(* IEC 61131-3 sources: plc-st-coding-agent/progress/evidence/f14_v5_public_pilot_20261112/jobs/codex_minimax-m27, 24 files *)

(* ---- public-easy-01.candidate_01.st ---- *)
(*
ENGINEERING_CONTRACT - Filling Line Control FB
==============================================
State Machine: Sequential, 6 states (IDLE→CLEANING→FILLING→CAPPING→PACKING→COMPLETED→IDLE)
---------------------------------------------------------------------------------
| State       | Activation         | Retention              | Reset/Deactivation            |
---------------------------------------------------------------------------------
| IDLE        | bottleSensor=TRUE  | Hold until bottle      | Deact on bottleSensor:=TRUE   |
| CLEANING    | cleaningConfirm    | Pump_Motor ON hold     | Deact on cleaningConfirm      |
| FILLING     | fillingConfirm     | Filling_Valve ON hold  | Deact on fillingConfirm       |
| CAPPING     | cappingConfirm     | Capping_Machine ON hold| Deact on cappingConfirm       |
| PACKING     | packingConfirm     | Packing_Machine ON hold| Deact on packingConfirm       |
| COMPLETED   | packingConfirm     | Completion_Light ON    | Deact on finishedButton       |
---------------------------------------------------------------------------------
Priority: IDLE > COMPLETED > CLEANING > FILLING > CAPPING > PACKING (same-scan)
Units: All inputs/outputs BOOL; all states enumerated; no TIME/LTIME used
Boundaries: bottleSensor triggers only from IDLE; finishedButton resets only from COMPLETED
PUB refs: PUB001, PUB003, PUB004, PUB005, PUB006, PUB007, PUB008
---------------------------------------------------------------------------------
*)
FUNCTION_BLOCK FillingLineControl
VAR
    eState : EFillState := EFillState.IDLE;
END_VAR

TYPE EFillState :
(
    IDLE       := 0,
    CLEANING   := 1,
    FILLING    := 2,
    CAPPING    := 3,
    PACKING    := 4,
    COMPLETED  := 5
);
END_TYPE;

CASE eState OF
    EFillState.IDLE:
        Pump_Motor       := FALSE;
        Filling_Valve    := FALSE;
        Capping_Machine  := FALSE;
        Packing_Machine  := FALSE;
        Completion_Light := FALSE;

        IF bottleSensor THEN
            eState := EFillState.CLEANING;
        END_IF;

    EFillState.CLEANING:
        Pump_Motor       := TRUE;
        Filling_Valve    := FALSE;
        Capping_Machine  := FALSE;
        Packing_Machine  := FALSE;
        Completion_Light := FALSE;

        IF cleaningConfirmButton THEN
            eState := EFillState.FILLING;
        END_IF;

    EFillState.FILLING:
        Pump_Motor       := TRUE;
        Filling_Valve    := TRUE;
        Capping_Machine  := FALSE;
        Packing_Machine  := FALSE;
        Completion_Light := FALSE;

        IF fillingConfirmButton THEN
            eState := EFillState.CAPPING;
        END_IF;

    EFillState.CAPPING:
        Pump_Motor       := TRUE;
        Filling_Valve    := FALSE;
        Capping_Machine  := TRUE;
        Packing_Machine  := FALSE;
        Completion_Light := FALSE;

        IF cappingConfirmButton THEN
            eState := EFillState.PACKING;
        END_IF;

    EFillState.PACKING:
        Pump_Motor       := TRUE;
        Filling_Valve    := FALSE;
        Capping_Machine  := FALSE;
        Packing_Machine  := TRUE;
        Completion_Light := FALSE;

        IF packingConfirmButton THEN
            eState := EFillState.COMPLETED;
        END_IF;

    EFillState.COMPLETED:
        Pump_Motor       := TRUE;
        Filling_Valve    := FALSE;
        Capping_Machine  := FALSE;
        Packing_Machine  := FALSE;
        Completion_Light := TRUE;

        IF finishedButton THEN
            eState := EFillState.IDLE;
        END_IF;

END_CASE;

END_FUNCTION_BLOCK

(* ---- public-easy-01.candidate_02.st ---- *)
(*
ENGINEERING_CONTRACT - Filling Line Control FB
==============================================
State Machine: Sequential, 6 states (IDLE→CLEANING→FILLING→CAPPING→PACKING→COMPLETED→IDLE)
---------------------------------------------------------------------------------
| State       | Activation         | Retention              | Reset/Deactivation            |
---------------------------------------------------------------------------------
| IDLE        | bottleSensor=TRUE  | Hold until bottle      | Deact on bottleSensor:=TRUE   |
| CLEANING    | cleaningConfirm    | Pump_Motor ON hold     | Deact on cleaningConfirm      |
| FILLING     | fillingConfirm     | Filling_Valve ON hold  | Deact on fillingConfirm       |
| CAPPING     | cappingConfirm     | Capping_Machine ON hold| Deact on cappingConfirm       |
| PACKING     | packingConfirm     | Packing_Machine ON hold| Deact on packingConfirm       |
| COMPLETED   | packingConfirm     | Completion_Light ON    | Deact on finishedButton       |
---------------------------------------------------------------------------------
Priority: IDLE > COMPLETED > CLEANING > FILLING > CAPPING > PACKING (same-scan)
Units: All inputs/outputs BOOL; all states enumerated; no TIME/LTIME used
Boundaries: bottleSensor triggers only from IDLE; finishedButton resets only from COMPLETED
PUB refs: PUB001, PUB003, PUB004, PUB005, PUB006, PUB007, PUB008
---------------------------------------------------------------------------------
*)
TYPE EFillState :
(
    IDLE       := 0,
    CLEANING   := 1,
    FILLING    := 2,
    CAPPING    := 3,
    PACKING    := 4,
    COMPLETED  := 5
);
END_TYPE;

FUNCTION_BLOCK FillingLineControl
VAR_INPUT
    bottleSensor           : BOOL;
    cleaningConfirmButton  : BOOL;
    fillingConfirmButton   : BOOL;
    cappingConfirmButton   : BOOL;
    packingConfirmButton   : BOOL;
    finishedButton         : BOOL;
END_VAR
VAR_OUTPUT
    Pump_Motor       : BOOL;
    Filling_Valve    : BOOL;
    Capping_Machine  : BOOL;
    Packing_Machine  : BOOL;
    Completion_Light : BOOL;
END_VAR
VAR
    eState : EFillState := EFillState.IDLE;
END_VAR

CASE eState OF
    EFillState.IDLE:
        Pump_Motor       := FALSE;
        Filling_Valve    := FALSE;
        Capping_Machine  := FALSE;
        Packing_Machine  := FALSE;
        Completion_Light := FALSE;

        IF bottleSensor THEN
            eState := EFillState.CLEANING;
        END_IF;

    EFillState.CLEANING:
        Pump_Motor       := TRUE;
        Filling_Valve    := FALSE;
        Capping_Machine  := FALSE;
        Packing_Machine  := FALSE;
        Completion_Light := FALSE;

        IF cleaningConfirmButton THEN
            eState := EFillState.FILLING;
        END_IF;

    EFillState.FILLING:
        Pump_Motor       := FALSE;
        Filling_Valve    := TRUE;
        Capping_Machine  := FALSE;
        Packing_Machine  := FALSE;
        Completion_Light := FALSE;

        IF fillingConfirmButton THEN
            eState := EFillState.CAPPING;
        END_IF;

    EFillState.CAPPING:
        Pump_Motor       := FALSE;
        Filling_Valve    := FALSE;
        Capping_Machine  := TRUE;
        Packing_Machine  := FALSE;
        Completion_Light := FALSE;

        IF cappingConfirmButton THEN
            eState := EFillState.PACKING;
        END_IF;

    EFillState.PACKING:
        Pump_Motor       := FALSE;
        Filling_Valve    := FALSE;
        Capping_Machine  := FALSE;
        Packing_Machine  := TRUE;
        Completion_Light := FALSE;

        IF packingConfirmButton THEN
            eState := EFillState.COMPLETED;
        END_IF;

    EFillState.COMPLETED:
        Pump_Motor       := FALSE;
        Filling_Valve    := FALSE;
        Capping_Machine  := FALSE;
        Packing_Machine  := FALSE;
        Completion_Light := TRUE;

        IF finishedButton THEN
            eState := EFillState.IDLE;
        END_IF;

END_CASE;

END_FUNCTION_BLOCK

(* ---- public-easy-01.raw_candidate_01.st ---- *)
(*
ENGINEERING_CONTRACT - Filling Line Control FB
==============================================
State Machine: Sequential, 6 states (IDLE→CLEANING→FILLING→CAPPING→PACKING→COMPLETED→IDLE)
---------------------------------------------------------------------------------
| State       | Activation         | Retention              | Reset/Deactivation            |
---------------------------------------------------------------------------------
| IDLE        | bottleSensor=TRUE  | Hold until bottle      | Deact on bottleSensor:=TRUE   |
| CLEANING    | cleaningConfirm    | Pump_Motor ON hold     | Deact on cleaningConfirm      |
| FILLING     | fillingConfirm     | Filling_Valve ON hold  | Deact on fillingConfirm       |
| CAPPING     | cappingConfirm     | Capping_Machine ON hold| Deact on cappingConfirm       |
| PACKING     | packingConfirm     | Packing_Machine ON hold| Deact on packingConfirm       |
| COMPLETED   | packingConfirm     | Completion_Light ON    | Deact on finishedButton       |
---------------------------------------------------------------------------------
Priority: IDLE > COMPLETED > CLEANING > FILLING > CAPPING > PACKING (same-scan)
Units: All inputs/outputs BOOL; all states enumerated; no TIME/LTIME used
Boundaries: bottleSensor triggers only from IDLE; finishedButton resets only from COMPLETED
PUB refs: PUB001, PUB003, PUB004, PUB005, PUB006, PUB007, PUB008
---------------------------------------------------------------------------------
*)
FUNCTION_BLOCK FillingLineControl
VAR
    eState : EFillState := EFillState.IDLE;
END_VAR

TYPE EFillState :
(
    IDLE       := 0,
    CLEANING   := 1,
    FILLING    := 2,
    CAPPING    := 3,
    PACKING    := 4,
    COMPLETED  := 5
);
END_TYPE

CASE eState OF
    EFillState.IDLE:
        Pump_Motor       := FALSE;
        Filling_Valve    := FALSE;
        Capping_Machine  := FALSE;
        Packing_Machine  := FALSE;
        Completion_Light := FALSE;

        IF bottleSensor THEN
            eState := EFillState.CLEANING;
        END_IF;

    EFillState.CLEANING:
        Pump_Motor       := TRUE;
        Filling_Valve    := FALSE;
        Capping_Machine  := FALSE;
        Packing_Machine  := FALSE;
        Completion_Light := FALSE;

        IF cleaningConfirmButton THEN
            eState := EFillState.FILLING;
        END_IF;

    EFillState.FILLING:
        Pump_Motor       := TRUE;
        Filling_Valve    := TRUE;
        Capping_Machine  := FALSE;
        Packing_Machine  := FALSE;
        Completion_Light := FALSE;

        IF fillingConfirmButton THEN
            eState := EFillState.CAPPING;
        END_IF;

    EFillState.CAPPING:
        Pump_Motor       := TRUE;
        Filling_Valve    := FALSE;
        Capping_Machine  := TRUE;
        Packing_Machine  := FALSE;
        Completion_Light := FALSE;

        IF cappingConfirmButton THEN
            eState := EFillState.PACKING;
        END_IF;

    EFillState.PACKING:
        Pump_Motor       := TRUE;
        Filling_Valve    := FALSE;
        Capping_Machine  := FALSE;
        Packing_Machine  := TRUE;
        Completion_Light := FALSE;

        IF packingConfirmButton THEN
            eState := EFillState.COMPLETED;
        END_IF;

    EFillState.COMPLETED:
        Pump_Motor       := TRUE;
        Filling_Valve    := FALSE;
        Capping_Machine  := FALSE;
        Packing_Machine  := FALSE;
        Completion_Light := TRUE;

        IF finishedButton THEN
            eState := EFillState.IDLE;
        END_IF;

END_CASE;

END_FUNCTION_BLOCK

(* ---- public-easy-01.raw_candidate_02.st ---- *)
(*
ENGINEERING_CONTRACT - Filling Line Control FB
==============================================
State Machine: Sequential, 6 states (IDLE→CLEANING→FILLING→CAPPING→PACKING→COMPLETED→IDLE)
---------------------------------------------------------------------------------
| State       | Activation         | Retention              | Reset/Deactivation            |
---------------------------------------------------------------------------------
| IDLE        | bottleSensor=TRUE  | Hold until bottle      | Deact on bottleSensor:=TRUE   |
| CLEANING    | cleaningConfirm    | Pump_Motor ON hold     | Deact on cleaningConfirm      |
| FILLING     | fillingConfirm     | Filling_Valve ON hold  | Deact on fillingConfirm       |
| CAPPING     | cappingConfirm     | Capping_Machine ON hold| Deact on cappingConfirm       |
| PACKING     | packingConfirm     | Packing_Machine ON hold| Deact on packingConfirm       |
| COMPLETED   | packingConfirm     | Completion_Light ON    | Deact on finishedButton       |
---------------------------------------------------------------------------------
Priority: IDLE > COMPLETED > CLEANING > FILLING > CAPPING > PACKING (same-scan)
Units: All inputs/outputs BOOL; all states enumerated; no TIME/LTIME used
Boundaries: bottleSensor triggers only from IDLE; finishedButton resets only from COMPLETED
PUB refs: PUB001, PUB003, PUB004, PUB005, PUB006, PUB007, PUB008
---------------------------------------------------------------------------------
*)
TYPE EFillState :
(
    IDLE       := 0,
    CLEANING   := 1,
    FILLING    := 2,
    CAPPING    := 3,
    PACKING    := 4,
    COMPLETED  := 5
);
END_TYPE

FUNCTION_BLOCK FillingLineControl
VAR_INPUT
    bottleSensor           : BOOL;
    cleaningConfirmButton  : BOOL;
    fillingConfirmButton   : BOOL;
    cappingConfirmButton   : BOOL;
    packingConfirmButton   : BOOL;
    finishedButton         : BOOL;
END_VAR
VAR_OUTPUT
    Pump_Motor       : BOOL;
    Filling_Valve    : BOOL;
    Capping_Machine  : BOOL;
    Packing_Machine  : BOOL;
    Completion_Light : BOOL;
END_VAR
VAR
    eState : EFillState := EFillState.IDLE;
END_VAR

CASE eState OF
    EFillState.IDLE:
        Pump_Motor       := FALSE;
        Filling_Valve    := FALSE;
        Capping_Machine  := FALSE;
        Packing_Machine  := FALSE;
        Completion_Light := FALSE;

        IF bottleSensor THEN
            eState := EFillState.CLEANING;
        END_IF;

    EFillState.CLEANING:
        Pump_Motor       := TRUE;
        Filling_Valve    := FALSE;
        Capping_Machine  := FALSE;
        Packing_Machine  := FALSE;
        Completion_Light := FALSE;

        IF cleaningConfirmButton THEN
            eState := EFillState.FILLING;
        END_IF;

    EFillState.FILLING:
        Pump_Motor       := FALSE;
        Filling_Valve    := TRUE;
        Capping_Machine  := FALSE;
        Packing_Machine  := FALSE;
        Completion_Light := FALSE;

        IF fillingConfirmButton THEN
            eState := EFillState.CAPPING;
        END_IF;

    EFillState.CAPPING:
        Pump_Motor       := FALSE;
        Filling_Valve    := FALSE;
        Capping_Machine  := TRUE;
        Packing_Machine  := FALSE;
        Completion_Light := FALSE;

        IF cappingConfirmButton THEN
            eState := EFillState.PACKING;
        END_IF;

    EFillState.PACKING:
        Pump_Motor       := FALSE;
        Filling_Valve    := FALSE;
        Capping_Machine  := FALSE;
        Packing_Machine  := TRUE;
        Completion_Light := FALSE;

        IF packingConfirmButton THEN
            eState := EFillState.COMPLETED;
        END_IF;

    EFillState.COMPLETED:
        Pump_Motor       := FALSE;
        Filling_Valve    := FALSE;
        Capping_Machine  := FALSE;
        Packing_Machine  := FALSE;
        Completion_Light := TRUE;

        IF finishedButton THEN
            eState := EFillState.IDLE;
        END_IF;

END_CASE;

END_FUNCTION_BLOCK

(* ---- public-easy-04.candidate_01.st ---- *)
FUNCTION_BLOCK JamPumpControl
VAR_INPUT
    VISCOSITY_OK    : BOOL;
    PASTE_E_STOP_NC : BOOL;
    DebounceTime    : TIME;
    CycleTime       : TIME;
END_VAR
VAR_OUTPUT
    VFD_RUN          : BOOL := FALSE;
    PUMP_MAINT_DUE   : BOOL := FALSE;
    PUMP_RUNTIME_ACC : LTIME := LTIME#0s;
END_VAR
VAR
    ViscosityDebounceTimer : TON;
    ViscosityDebounceAccum : LTIME := LTIME#0s;
    ViscosityValid         : BOOL := FALSE;
END_VAR
// ENGINEERING_CONTRACT
// | Output/State    | Activation         | Retention          | Reset/Deactivation                      | Priority | Units/Boundaries |
// |-----------------|--------------------|--------------------|-----------------------------------------|----------|-------------------|
// | VFD_RUN         | TRUE when safety   | Retained while     | Cleared on E-Stop or viscosity invalid  | Safety   | Boolean permissive|
// |                 | permissive AND     | conditions met     | (PUB003)                                | first    |                   |
// |                 | viscosity valid    |                    |                                         |          |                   |
// | PUMP_MAINT_DUE  | Set when runtime   | Latched TRUE       | No reset (informational only, PUB004)   | None     | 500h threshold    |
// |                 | >= 500h (PUB004)   |                    |                                         |          |                   |
// | PUMP_RUNTIME_ACC| Increments by      | Preserved when     | Init to 0 at power-up only (PUB005)     | None     | LTIME (nanoseconds)|
// |                 | CycleTime when     | VFD_RUN = FALSE    |                                         |          | 0 to max          |
// |                 | VFD_RUN = TRUE     | (PUB003)           |                                         |          |                   |
// |                 | (PUB003)          |                    |                                         |          |                   |
// | ViscosityValid  | After DebounceTime | Retained while     | Immediate on VISCITY_OK=FALSE or        | None     | Debounced state   |
// |                 | continuous TRUE    | VISCOSITY_OK=TRUE  | E-Stop (PUB002, PUB003)                 |          |                   |
// |                 | (PUB002)          | (PUB002)           |                                         |          |                   |
// | ViscosityDebounceAccum | Accumulates  | Reset to 0 when   | Reset on VISCOSITY_OK=FALSE or          | None     | LTIME nanoseconds |
// |                 | elapsed time when  | VISCOSITY_OK=FALSE | E-Stop (PUB003)                         |          | >= 0              |
// |                 | VISCOSITY_OK=TRUE  |                    |                                         |          |                   |

// Viscosity debouncing (PUB002)
IF NOT VISCOSITY_OK THEN
    ViscosityDebounceAccum := LTIME#0s;
    ViscosityValid := FALSE;
    ViscosityDebounceTimer(IN := FALSE);
ELSIF ViscosityValid THEN
    ViscosityDebounceTimer(IN := TRUE, PT := DebounceTime);
ELSE
    ViscosityDebounceAccum := ViscosityDebounceAccum + CycleTime;
    IF ViscosityDebounceAccum >= DebounceTime THEN
        ViscosityValid := TRUE;
    END_IF;
    ViscosityDebounceTimer(IN := FALSE);
END_IF;

// Safety permissive and run command (PUB003)
IF NOT PASTE_E_STOP_NC THEN
    VFD_RUN := FALSE;
    ViscosityDebounceAccum := LTIME#0s;
    ViscosityValid := FALSE;
END_IF;

IF PASTE_E_STOP_NC AND ViscosityValid THEN
    VFD_RUN := TRUE;
ELSE
    VFD_RUN := FALSE;
END_IF;

// Runtime accumulation (PUB003, PUB004)
IF VFD_RUN THEN
    PUMP_RUNTIME_ACC := PUMP_RUNTIME_ACC + CycleTime;
END_IF;

IF PUMP_RUNTIME_ACC >= T#500h THEN
    PUMP_MAINT_DUE := TRUE;
END_IF;
END_FUNCTION_BLOCK

(* ---- public-easy-04.candidate_02.st ---- *)
FUNCTION_BLOCK JamPumpControl
VAR_INPUT
    VISCOSITY_OK    : BOOL;
    PASTE_E_STOP_NC : BOOL;
    DebounceTime    : TIME;
    CycleTime       : TIME;
END_VAR
VAR_OUTPUT
    VFD_RUN          : BOOL := FALSE;
    PUMP_MAINT_DUE   : BOOL := FALSE;
    PUMP_RUNTIME_ACC : LTIME := LTIME#0s;
END_VAR
VAR
    ViscosityValid         : BOOL := FALSE;
    ViscosityDebounceAccum : LTIME := LTIME#0s;
    DebounceTarget         : LTIME;
    CycleAsLTIME           : LTIME;
END_VAR
// ENGINEERING_CONTRACT
// | Output/State             | Activation                          | Retention            | Reset/Deactivation                      | Priority | Units/Boundaries |
// |--------------------------|-------------------------------------|----------------------|-----------------------------------------|----------|-------------------|
// | VFD_RUN                  | TRUE when safety permissive AND     | Retained while       | Cleared on E-Stop or viscosity invalid  | Safety   | Boolean permissive|
// |                          | viscosity valid (PUB003)            | conditions met       | (PUB003)                                | first    |                   |
// | PUMP_MAINT_DUE           | Set when runtime >= 500h (PUB004)   | Latched TRUE         | No reset (informational only, PUB004)   | None     | 500h threshold    |
// | PUMP_RUNTIME_ACC         | Increments by CycleTime when        | Preserved when       | Init to 0 at power-up only (PUB005)     | None     | LTIME nanoseconds |
// |                          | VFD_RUN = TRUE (PUB003)             | VFD_RUN = FALSE      |                                         |          | 0 to max          |
// | ViscosityValid           | After DebounceTime continuous TRUE  | Retained while       | Immediate on VISCOSITY_OK=FALSE or      | None     | Debounced state   |
// |                          | (PUB002)                            | VISCITY_OK=TRUE      | E-Stop (PUB002, PUB003)                 |          |                   |
// | ViscosityDebounceAccum   | Accumulates elapsed time when       | Reset to 0 when      | Reset on VISCOSITY_OK=FALSE or          | None     | LTIME nanoseconds |
// |                          | VISCOSITY_OK=TRUE (PUB002)          | VISCITY_OK=FALSE     | E-Stop (PUB003)                         |          | >= 0              |

DebounceTarget := TIME_TO_LTIME(DebounceTime);
CycleAsLTIME   := TIME_TO_LTIME(CycleTime);

// Emergency stop immediately clears run output and debounce state (PUB003)
IF NOT PASTE_E_STOP_NC THEN
    VFD_RUN := FALSE;
    ViscosityDebounceAccum := LTIME#0s;
    ViscosityValid := FALSE;
END_IF;

// Viscosity debouncing (PUB002): invalidate immediately on FALSE
IF NOT VISCOSITY_OK THEN
    ViscosityDebounceAccum := LTIME#0s;
    ViscosityValid := FALSE;
ELSE
    // Accumulate only when viscosity TRUE and not yet valid
    IF NOT ViscosityValid THEN
        ViscosityDebounceAccum := ViscosityDebounceAccum + CycleAsLTIME;
        IF ViscosityDebounceAccum >= DebounceTarget THEN
            ViscosityValid := TRUE;
        END_IF;
    END_IF;
END_IF;

// VFD_RUN permissive (PUB003)
IF PASTE_E_STOP_NC AND ViscosityValid THEN
    VFD_RUN := TRUE;
ELSE
    VFD_RUN := FALSE;
END_IF;

// Runtime accumulation (PUB003, PUB004)
IF VFD_RUN THEN
    PUMP_RUNTIME_ACC := PUMP_RUNTIME_ACC + CycleAsLTIME;
END_IF;

IF PUMP_RUNTIME_ACC >= LTIME#500h THEN
    PUMP_MAINT_DUE := TRUE;
END_IF;
END_FUNCTION_BLOCK

(* ---- public-easy-04.raw_candidate_01.st ---- *)
FUNCTION_BLOCK JamPumpControl
VAR_INPUT
    VISCOSITY_OK    : BOOL;
    PASTE_E_STOP_NC : BOOL;
    DebounceTime    : TIME;
    CycleTime       : TIME;
END_VAR
VAR_OUTPUT
    VFD_RUN          : BOOL := FALSE;
    PUMP_MAINT_DUE   : BOOL := FALSE;
    PUMP_RUNTIME_ACC : LTIME := LTIME#0s;
END_VAR
VAR
    ViscosityDebounceTimer : TON;
    ViscosityDebounceAccum : LTIME := LTIME#0s;
    ViscosityValid         : BOOL := FALSE;
END_VAR
// ENGINEERING_CONTRACT
// | Output/State    | Activation         | Retention          | Reset/Deactivation                      | Priority | Units/Boundaries |
// |-----------------|--------------------|--------------------|-----------------------------------------|----------|-------------------|
// | VFD_RUN         | TRUE when safety   | Retained while     | Cleared on E-Stop or viscosity invalid  | Safety   | Boolean permissive|
// |                 | permissive AND     | conditions met     | (PUB003)                                | first    |                   |
// |                 | viscosity valid    |                    |                                         |          |                   |
// | PUMP_MAINT_DUE  | Set when runtime   | Latched TRUE       | No reset (informational only, PUB004)   | None     | 500h threshold    |
// |                 | >= 500h (PUB004)   |                    |                                         |          |                   |
// | PUMP_RUNTIME_ACC| Increments by      | Preserved when     | Init to 0 at power-up only (PUB005)     | None     | LTIME (nanoseconds)|
// |                 | CycleTime when     | VFD_RUN = FALSE    |                                         |          | 0 to max          |
// |                 | VFD_RUN = TRUE     | (PUB003)           |                                         |          |                   |
// |                 | (PUB003)          |                    |                                         |          |                   |
// | ViscosityValid  | After DebounceTime | Retained while     | Immediate on VISCITY_OK=FALSE or        | None     | Debounced state   |
// |                 | continuous TRUE    | VISCOSITY_OK=TRUE  | E-Stop (PUB002, PUB003)                 |          |                   |
// |                 | (PUB002)          | (PUB002)           |                                         |          |                   |
// | ViscosityDebounceAccum | Accumulates  | Reset to 0 when   | Reset on VISCOSITY_OK=FALSE or          | None     | LTIME nanoseconds |
// |                 | elapsed time when  | VISCOSITY_OK=FALSE | E-Stop (PUB003)                         |          | >= 0              |
// |                 | VISCOSITY_OK=TRUE  |                    |                                         |          |                   |

// Viscosity debouncing (PUB002)
IF NOT VISCOSITY_OK THEN
    ViscosityDebounceAccum := LTIME#0s;
    ViscosityValid := FALSE;
    ViscosityDebounceTimer(IN := FALSE);
ELSIF ViscosityValid THEN
    ViscosityDebounceTimer(IN := TRUE, PT := DebounceTime);
ELSE
    ViscosityDebounceAccum := ViscosityDebounceAccum + CycleTime;
    IF ViscosityDebounceAccum >= DebounceTime THEN
        ViscosityValid := TRUE;
    END_IF
    ViscosityDebounceTimer(IN := FALSE);
END_IF;

// Safety permissive and run command (PUB003)
IF NOT PASTE_E_STOP_NC THEN
    VFD_RUN := FALSE;
    ViscosityDebounceAccum := LTIME#0s;
    ViscosityValid := FALSE;
END_IF;

IF PASTE_E_STOP_NC AND ViscosityValid THEN
    VFD_RUN := TRUE;
ELSE
    VFD_RUN := FALSE;
END_IF;

// Runtime accumulation (PUB003, PUB004)
IF VFD_RUN THEN
    PUMP_RUNTIME_ACC := PUMP_RUNTIME_ACC + CycleTime;
END_IF;

IF PUMP_RUNTIME_ACC >= T#500h THEN
    PUMP_MAINT_DUE := TRUE;
END_IF;
END_FUNCTION_BLOCK

(* ---- public-easy-04.raw_candidate_02.st ---- *)
FUNCTION_BLOCK JamPumpControl
VAR_INPUT
    VISCOSITY_OK    : BOOL;
    PASTE_E_STOP_NC : BOOL;
    DebounceTime    : TIME;
    CycleTime       : TIME;
END_VAR
VAR_OUTPUT
    VFD_RUN          : BOOL := FALSE;
    PUMP_MAINT_DUE   : BOOL := FALSE;
    PUMP_RUNTIME_ACC : LTIME := LTIME#0s;
END_VAR
VAR
    ViscosityValid         : BOOL := FALSE;
    ViscosityDebounceAccum : LTIME := LTIME#0s;
    DebounceTarget         : LTIME;
    CycleAsLTIME           : LTIME;
END_VAR
// ENGINEERING_CONTRACT
// | Output/State             | Activation                          | Retention            | Reset/Deactivation                      | Priority | Units/Boundaries |
// |--------------------------|-------------------------------------|----------------------|-----------------------------------------|----------|-------------------|
// | VFD_RUN                  | TRUE when safety permissive AND     | Retained while       | Cleared on E-Stop or viscosity invalid  | Safety   | Boolean permissive|
// |                          | viscosity valid (PUB003)            | conditions met       | (PUB003)                                | first    |                   |
// | PUMP_MAINT_DUE           | Set when runtime >= 500h (PUB004)   | Latched TRUE         | No reset (informational only, PUB004)   | None     | 500h threshold    |
// | PUMP_RUNTIME_ACC         | Increments by CycleTime when        | Preserved when       | Init to 0 at power-up only (PUB005)     | None     | LTIME nanoseconds |
// |                          | VFD_RUN = TRUE (PUB003)             | VFD_RUN = FALSE      |                                         |          | 0 to max          |
// | ViscosityValid           | After DebounceTime continuous TRUE  | Retained while       | Immediate on VISCOSITY_OK=FALSE or      | None     | Debounced state   |
// |                          | (PUB002)                            | VISCITY_OK=TRUE      | E-Stop (PUB002, PUB003)                 |          |                   |
// | ViscosityDebounceAccum   | Accumulates elapsed time when       | Reset to 0 when      | Reset on VISCOSITY_OK=FALSE or          | None     | LTIME nanoseconds |
// |                          | VISCOSITY_OK=TRUE (PUB002)          | VISCITY_OK=FALSE     | E-Stop (PUB003)                         |          | >= 0              |

DebounceTarget := TIME_TO_LTIME(DebounceTime);
CycleAsLTIME   := TIME_TO_LTIME(CycleTime);

// Emergency stop immediately clears run output and debounce state (PUB003)
IF NOT PASTE_E_STOP_NC THEN
    VFD_RUN := FALSE;
    ViscosityDebounceAccum := LTIME#0s;
    ViscosityValid := FALSE;
END_IF;

// Viscosity debouncing (PUB002): invalidate immediately on FALSE
IF NOT VISCOSITY_OK THEN
    ViscosityDebounceAccum := LTIME#0s;
    ViscosityValid := FALSE;
ELSE
    // Accumulate only when viscosity TRUE and not yet valid
    IF NOT ViscosityValid THEN
        ViscosityDebounceAccum := ViscosityDebounceAccum + CycleAsLTIME;
        IF ViscosityDebounceAccum >= DebounceTarget THEN
            ViscosityValid := TRUE;
        END_IF;
    END_IF;
END_IF;

// VFD_RUN permissive (PUB003)
IF PASTE_E_STOP_NC AND ViscosityValid THEN
    VFD_RUN := TRUE;
ELSE
    VFD_RUN := FALSE;
END_IF;

// Runtime accumulation (PUB003, PUB004)
IF VFD_RUN THEN
    PUMP_RUNTIME_ACC := PUMP_RUNTIME_ACC + CycleAsLTIME;
END_IF;

IF PUMP_RUNTIME_ACC >= LTIME#500h THEN
    PUMP_MAINT_DUE := TRUE;
END_IF;
END_FUNCTION_BLOCK

(* ---- public-hard-03.candidate_01.st ---- *)
(* ENGINEERING_CONTRACT: Recipe Management System FB_RecipeManager
+------------------------------------------------------------------
| PUB001-006: CRUD operations on recipe database (ARRAY[1..10])
| Output State Groups:
|   - recipeAdded/Deleted/Modified: activation on success, reset
|     when input goes FALSE (level-triggered, same-scan)
|   - recipeQueryResult: populated on success (no separate success flag)
|   - error+status: activation on failure, reset on success
| Priority: Sequential IF chain; query > add > delete > modify
| Units: recipeID(INT), ingredientType(INT), ingredientRatio(REAL),
|        productionTemperature(REAL)
| Boundaries: recipeID=0 denotes empty slot; array bounds 1..10
+------------------------------------------------------------------ *)

TYPE ST_Recipe : STRUCT
    recipeID             : INT;
    ingredientType       : INT;
    ingredientRatio      : REAL;
    productionTemperature: REAL;
END_STRUCT
END_TYPE;

FUNCTION_BLOCK FB_RecipeManager
VAR_INPUT
    addRecipe    : BOOL;
    deleteRecipe : BOOL;
    modifyRecipe : BOOL;
    queryRecipe  : BOOL;
    recipeIn     : ST_Recipe;
END_VAR
VAR_OUTPUT
    recipeAdded       : BOOL := FALSE;
    recipeDeleted     : BOOL := FALSE;
    recipeModified    : BOOL := FALSE;
    recipeQueryResult : ST_Recipe;
    error             : BOOL := FALSE;
    status            : WORD := 16#0000;
END_VAR
VAR_IN_OUT
    recipe : ARRAY[1..10] OF ST_Recipe;
END_VAR
VAR
    idx     : INT;
    found   : BOOL;
    emptyIdx: INT;
END_VAR

// Initialize per scan
error             := FALSE;
status            := 16#0000;
recipeAdded       := FALSE;
recipeDeleted     := FALSE;
recipeModified    := FALSE;
recipeQueryResult.recipeID             := 0;
recipeQueryResult.ingredientType       := 0;
recipeQueryResult.ingredientRatio      := 0.0;
recipeQueryResult.productionTemperature:= 0.0;

// PUB009: Query by recipeID
IF queryRecipe THEN
    found := FALSE;
    FOR idx := 1 TO 10 DO
        IF recipe[idx].recipeID = recipeIn.recipeID THEN
            recipeQueryResult := recipe[idx];
            found := TRUE;
            EXIT;
        END_IF;
    END_FOR;
    IF NOT found THEN
        error := TRUE;
        status := 16#8001;
    END_IF;
END_IF;

// PUB010: Add new recipe
IF addRecipe THEN
    found := FALSE;
    FOR idx := 1 TO 10 DO
        IF recipe[idx].recipeID = recipeIn.recipeID THEN
            found := TRUE;
            EXIT;
        END_IF;
    END_FOR;
    IF found THEN
        error := TRUE;
        status := 16#8002;
    ELSE
        emptyIdx := 0;
        FOR idx := 1 TO 10 DO
            IF recipe[idx].recipeID = 0 THEN
                emptyIdx := idx;
                EXIT;
            END_IF;
        END_FOR;
        IF emptyIdx = 0 THEN
            error := TRUE;
            status := 16#8003;
        ELSE
            recipe[emptyIdx] := recipeIn;
            recipeAdded := TRUE;
        END_IF;
    END_IF;
END_IF;

// PUB011: Delete recipe by setting recipeID to 0
IF deleteRecipe THEN
    found := FALSE;
    FOR idx := 1 TO 10 DO
        IF recipe[idx].recipeID = recipeIn.recipeID THEN
            recipe[idx].recipeID := 0;
            found := TRUE;
            EXIT;
        END_IF;
    END_FOR;
    IF NOT found THEN
        error := TRUE;
        status := 16#8004;
    ELSE
        recipeDeleted := TRUE;
    END_IF;
END_IF;

// PUB012: Modify existing recipe
IF modifyRecipe THEN
    found := FALSE;
    FOR idx := 1 TO 10 DO
        IF recipe[idx].recipeID = recipeIn.recipeID THEN
            recipe[idx] := recipeIn;
            found := TRUE;
            EXIT;
        END_IF;
    END_FOR;
    IF NOT found THEN
        error := TRUE;
        status := 16#8005;
    ELSE
        recipeModified := TRUE;
    END_IF;
END_IF;
END_FUNCTION_BLOCK

(* ---- public-hard-03.candidate_02.st ---- *)
(* ENGINEERING_CONTRACT: Recipe Management System FB_RecipeManager
+------------------------------------------------------------------
| PUB001-006: CRUD operations on recipe database (ARRAY[1..10])
| Output State Groups:
|   - recipeAdded/Deleted/Modified: activation on success, reset
|     when input goes FALSE (level-triggered, same-scan)
|   - recipeQueryResult: populated on success (no separate success flag)
|   - error+status: activation on failure, reset on success
| Priority: Sequential IF chain; query > add > delete > modify
| Units: recipeID(INT), ingredientType(INT), ingredientRatio(REAL),
|        productionTemperature(REAL)
| Boundaries: recipeID=0 denotes empty slot; array bounds 1..10
+------------------------------------------------------------------ *)

TYPE ST_Recipe : STRUCT
    recipeID             : INT;
    ingredientType       : INT;
    ingredientRatio      : REAL;
    productionTemperature: REAL;
END_STRUCT
END_TYPE;

FUNCTION_BLOCK FB_RecipeManager
VAR_INPUT
    addRecipe    : BOOL;
    deleteRecipe : BOOL;
    modifyRecipe : BOOL;
    queryRecipe  : BOOL;
    recipeIn     : ST_Recipe;
END_VAR
VAR_OUTPUT
    recipeAdded       : BOOL := FALSE;
    recipeDeleted     : BOOL := FALSE;
    recipeModified    : BOOL := FALSE;
    recipeQueryResult : ST_Recipe;
    error             : BOOL := FALSE;
    status            : WORD := 16#0000;
END_VAR
VAR_IN_OUT
    recipe : ARRAY[1..10] OF ST_Recipe;
END_VAR
VAR
    idx       : INT;
    found     : BOOL;
    emptySlot : INT;
END_VAR

// Reset outputs at start of each scan cycle
error             := FALSE;
status            := 16#0000;
recipeAdded       := FALSE;
recipeDeleted     := FALSE;
recipeModified    := FALSE;
recipeQueryResult.recipeID             := 0;
recipeQueryResult.ingredientType       := 0;
recipeQueryResult.ingredientRatio      := 0.0;
recipeQueryResult.productionTemperature:= 0.0;

// Initialize local state
found     := FALSE;
emptySlot := 0;

// PUB009: Query recipe by recipeID
IF queryRecipe THEN
    found := FALSE;
    FOR idx := 1 TO 10 DO
        IF recipe[idx].recipeID = recipeIn.recipeID THEN
            recipeQueryResult := recipe[idx];
            found := TRUE;
            EXIT;
        END_IF;
    END_FOR;
    IF NOT found THEN
        error := TRUE;
        status := 16#8001;
    END_IF;
END_IF;

// PUB010: Add new recipe
IF addRecipe THEN
    // Check for duplicate recipeID
    found := FALSE;
    FOR idx := 1 TO 10 DO
        IF recipe[idx].recipeID = recipeIn.recipeID THEN
            found := TRUE;
            EXIT;
        END_IF;
    END_FOR;

    IF found THEN
        error := TRUE;
        status := 16#8002;
    ELSE
        // Find first empty slot (smallest index)
        emptySlot := 0;
        FOR idx := 1 TO 10 DO
            IF recipe[idx].recipeID = 0 THEN
                emptySlot := idx;
                EXIT;
            END_IF;
        END_FOR;

        IF emptySlot = 0 THEN
            error := TRUE;
            status := 16#8003;
        ELSE
            recipe[emptySlot].recipeID              := recipeIn.recipeID;
            recipe[emptySlot].ingredientType        := recipeIn.ingredientType;
            recipe[emptySlot].ingredientRatio       := recipeIn.ingredientRatio;
            recipe[emptySlot].productionTemperature := recipeIn.productionTemperature;
            recipeAdded := TRUE;
        END_IF;
    END_IF;
END_IF;

// PUB011: Delete recipe by setting recipeID to 0
IF deleteRecipe THEN
    found := FALSE;
    FOR idx := 1 TO 10 DO
        IF recipe[idx].recipeID = recipeIn.recipeID THEN
            recipe[idx].recipeID := 0;
            recipeDeleted := TRUE;
            found := TRUE;
            EXIT;
        END_IF;
    END_FOR;

    IF NOT found THEN
        error := TRUE;
        status := 16#8004;
    END_IF;
END_IF;

// PUB012: Modify existing recipe
IF modifyRecipe THEN
    found := FALSE;
    FOR idx := 1 TO 10 DO
        IF recipe[idx].recipeID = recipeIn.recipeID THEN
            recipe[idx].recipeID              := recipeIn.recipeID;
            recipe[idx].ingredientType        := recipeIn.ingredientType;
            recipe[idx].ingredientRatio       := recipeIn.ingredientRatio;
            recipe[idx].productionTemperature := recipeIn.productionTemperature;
            recipeModified := TRUE;
            found := TRUE;
            EXIT;
        END_IF;
    END_FOR;

    IF NOT found THEN
        error := TRUE;
        status := 16#8005;
    END_IF;
END_IF;
END_FUNCTION_BLOCK

(* ---- public-hard-03.raw_candidate_01.st ---- *)
(* ENGINEERING_CONTRACT: Recipe Management System FB_RecipeManager
+------------------------------------------------------------------
| PUB001-006: CRUD operations on recipe database (ARRAY[1..10])
| Output State Groups:
|   - recipeAdded/Deleted/Modified: activation on success, reset
|     when input goes FALSE (level-triggered, same-scan)
|   - recipeQueryResult: populated on success (no separate success flag)
|   - error+status: activation on failure, reset on success
| Priority: Sequential IF chain; query > add > delete > modify
| Units: recipeID(INT), ingredientType(INT), ingredientRatio(REAL),
|        productionTemperature(REAL)
| Boundaries: recipeID=0 denotes empty slot; array bounds 1..10
+------------------------------------------------------------------ *)

TYPE ST_Recipe : STRUCT
    recipeID             : INT;
    ingredientType       : INT;
    ingredientRatio      : REAL;
    productionTemperature: REAL;
END_STRUCT
END_TYPE

FUNCTION_BLOCK FB_RecipeManager
VAR_INPUT
    addRecipe    : BOOL;
    deleteRecipe : BOOL;
    modifyRecipe : BOOL;
    queryRecipe  : BOOL;
    recipeIn     : ST_Recipe;
END_VAR
VAR_OUTPUT
    recipeAdded       : BOOL := FALSE;
    recipeDeleted     : BOOL := FALSE;
    recipeModified    : BOOL := FALSE;
    recipeQueryResult : ST_Recipe;
    error             : BOOL := FALSE;
    status            : WORD := 16#0000;
END_VAR
VAR_IN_OUT
    recipe : ARRAY[1..10] OF ST_Recipe;
END_VAR
VAR
    idx     : INT;
    found   : BOOL;
    emptyIdx: INT;
END_VAR

// Initialize per scan
error             := FALSE;
status            := 16#0000;
recipeAdded       := FALSE;
recipeDeleted     := FALSE;
recipeModified    := FALSE;
recipeQueryResult.recipeID             := 0;
recipeQueryResult.ingredientType       := 0;
recipeQueryResult.ingredientRatio      := 0.0;
recipeQueryResult.productionTemperature:= 0.0;

// PUB009: Query by recipeID
IF queryRecipe THEN
    found := FALSE;
    FOR idx := 1 TO 10 DO
        IF recipe[idx].recipeID = recipeIn.recipeID THEN
            recipeQueryResult := recipe[idx];
            found := TRUE;
            EXIT;
        END_IF
    END_FOR;
    IF NOT found THEN
        error := TRUE;
        status := 16#8001;
    END_IF;
END_IF;

// PUB010: Add new recipe
IF addRecipe THEN
    found := FALSE;
    FOR idx := 1 TO 10 DO
        IF recipe[idx].recipeID = recipeIn.recipeID THEN
            found := TRUE;
            EXIT;
        END_IF;
    END_FOR;
    IF found THEN
        error := TRUE;
        status := 16#8002;
    ELSE
        emptyIdx := 0;
        FOR idx := 1 TO 10 DO
            IF recipe[idx].recipeID = 0 THEN
                emptyIdx := idx;
                EXIT;
            END_IF;
        END_FOR;
        IF emptyIdx = 0 THEN
            error := TRUE;
            status := 16#8003;
        ELSE
            recipe[emptyIdx] := recipeIn;
            recipeAdded := TRUE;
        END_IF;
    END_IF;
END_IF;

// PUB011: Delete recipe by setting recipeID to 0
IF deleteRecipe THEN
    found := FALSE;
    FOR idx := 1 TO 10 DO
        IF recipe[idx].recipeID = recipeIn.recipeID THEN
            recipe[idx].recipeID := 0;
            found := TRUE;
            EXIT;
        END_IF;
    END_FOR;
    IF NOT found THEN
        error := TRUE;
        status := 16#8004;
    ELSE
        recipeDeleted := TRUE;
    END_IF;
END_IF;

// PUB012: Modify existing recipe
IF modifyRecipe THEN
    found := FALSE;
    FOR idx := 1 TO 10 DO
        IF recipe[idx].recipeID = recipeIn.recipeID THEN
            recipe[idx] := recipeIn;
            found := TRUE;
            EXIT;
        END_IF;
    END_FOR;
    IF NOT found THEN
        error := TRUE;
        status := 16#8005;
    ELSE
        recipeModified := TRUE;
    END_IF;
END_IF;
END_FUNCTION_BLOCK

(* ---- public-hard-03.raw_candidate_02.st ---- *)
(* ENGINEERING_CONTRACT: Recipe Management System FB_RecipeManager
+------------------------------------------------------------------
| PUB001-006: CRUD operations on recipe database (ARRAY[1..10])
| Output State Groups:
|   - recipeAdded/Deleted/Modified: activation on success, reset
|     when input goes FALSE (level-triggered, same-scan)
|   - recipeQueryResult: populated on success (no separate success flag)
|   - error+status: activation on failure, reset on success
| Priority: Sequential IF chain; query > add > delete > modify
| Units: recipeID(INT), ingredientType(INT), ingredientRatio(REAL),
|        productionTemperature(REAL)
| Boundaries: recipeID=0 denotes empty slot; array bounds 1..10
+------------------------------------------------------------------ *)

TYPE ST_Recipe : STRUCT
    recipeID             : INT;
    ingredientType       : INT;
    ingredientRatio      : REAL;
    productionTemperature: REAL;
END_STRUCT
END_TYPE;

FUNCTION_BLOCK FB_RecipeManager
VAR_INPUT
    addRecipe    : BOOL;
    deleteRecipe : BOOL;
    modifyRecipe : BOOL;
    queryRecipe  : BOOL;
    recipeIn     : ST_Recipe;
END_VAR
VAR_OUTPUT
    recipeAdded       : BOOL := FALSE;
    recipeDeleted     : BOOL := FALSE;
    recipeModified    : BOOL := FALSE;
    recipeQueryResult : ST_Recipe;
    error             : BOOL := FALSE;
    status            : WORD := 16#0000;
END_VAR
VAR_IN_OUT
    recipe : ARRAY[1..10] OF ST_Recipe;
END_VAR
VAR
    idx       : INT;
    found     : BOOL;
    emptySlot : INT;
END_VAR

// Reset outputs at start of each scan cycle
error             := FALSE;
status            := 16#0000;
recipeAdded       := FALSE;
recipeDeleted     := FALSE;
recipeModified    := FALSE;
recipeQueryResult.recipeID             := 0;
recipeQueryResult.ingredientType       := 0;
recipeQueryResult.ingredientRatio      := 0.0;
recipeQueryResult.productionTemperature:= 0.0;

// Initialize local state
found     := FALSE;
emptySlot := 0;

// PUB009: Query recipe by recipeID
IF queryRecipe THEN
    found := FALSE;
    FOR idx := 1 TO 10 DO
        IF recipe[idx].recipeID = recipeIn.recipeID THEN
            recipeQueryResult := recipe[idx];
            found := TRUE;
            EXIT;
        END_IF;
    END_FOR;
    IF NOT found THEN
        error := TRUE;
        status := 16#8001;
    END_IF;
END_IF;

// PUB010: Add new recipe
IF addRecipe THEN
    // Check for duplicate recipeID
    found := FALSE;
    FOR idx := 1 TO 10 DO
        IF recipe[idx].recipeID = recipeIn.recipeID THEN
            found := TRUE;
            EXIT;
        END_IF;
    END_FOR;

    IF found THEN
        error := TRUE;
        status := 16#8002;
    ELSE
        // Find first empty slot (smallest index)
        emptySlot := 0;
        FOR idx := 1 TO 10 DO
            IF recipe[idx].recipeID = 0 THEN
                emptySlot := idx;
                EXIT;
            END_IF;
        END_FOR;

        IF emptySlot = 0 THEN
            error := TRUE;
            status := 16#8003;
        ELSE
            recipe[emptySlot].recipeID              := recipeIn.recipeID;
            recipe[emptySlot].ingredientType        := recipeIn.ingredientType;
            recipe[emptySlot].ingredientRatio       := recipeIn.ingredientRatio;
            recipe[emptySlot].productionTemperature := recipeIn.productionTemperature;
            recipeAdded := TRUE;
        END_IF;
    END_IF;
END_IF;

// PUB011: Delete recipe by setting recipeID to 0
IF deleteRecipe THEN
    found := FALSE;
    FOR idx := 1 TO 10 DO
        IF recipe[idx].recipeID = recipeIn.recipeID THEN
            recipe[idx].recipeID := 0;
            recipeDeleted := TRUE;
            found := TRUE;
            EXIT;
        END_IF;
    END_FOR;

    IF NOT found THEN
        error := TRUE;
        status := 16#8004;
    END_IF;
END_IF;

// PUB012: Modify existing recipe
IF modifyRecipe THEN
    found := FALSE;
    FOR idx := 1 TO 10 DO
        IF recipe[idx].recipeID = recipeIn.recipeID THEN
            recipe[idx].recipeID              := recipeIn.recipeID;
            recipe[idx].ingredientType        := recipeIn.ingredientType;
            recipe[idx].ingredientRatio       := recipeIn.ingredientRatio;
            recipe[idx].productionTemperature := recipeIn.productionTemperature;
            recipeModified := TRUE;
            found := TRUE;
            EXIT;
        END_IF;
    END_FOR;

    IF NOT found THEN
        error := TRUE;
        status := 16#8005;
    END_IF;
END_IF;
END_FUNCTION_BLOCK

(* ---- public-medium-03.candidate_01.st ---- *)
FUNCTION_BLOCK FB_MovingAverage
(* Engineering Contract
 * ┌─────────────────────────────────────────────────────────────────────────────────────┐
 * │ OUTPUT STATE TABLE                                                                │
 * ├─────────────┬────────────────────────────────────────────────────────────────────┤
 * │ average     │ HOLD: Retained between scans; updated when valid sample processed.  │
 * │             │ RETAIN on reset: Returns to 0.0 via sum reset.                      │
 * │ windowSizeReached│ ACTIVE: TRUE when sampleCount >= windowSize (PUB001 window).   │
 * │             │ DEACTIVATION: Set FALSE on reset.                                   │
 * │ error       │ ACTIVE: TRUE when windowSize invalid (<1 or >100).                  │
 * │             │ DEACTIVATION: Set FALSE when reset clears error.                    │
 * │ status      │ RETAIN: 16#8200 when invalid windowSize; 16#0000 otherwise.         │
 * │             │ RESET: Set to 16#0000 on valid reset or valid windowSize.           │
 * ├─────────────┼────────────────────────────────────────────────────────────────────┤
 * │ TRIGGER     │ Rising edge on trigger input (PUB003). Edge detection via           │
 * │             │ triggerPrev state variable. Same-scan priority: cyclicExecution     │
 * │             │ checked first per PUB002.                                           │
 * ├─────────────┼────────────────────────────────────────────────────────────────────┤
 * │ WINDOW      │ Bounded 1..100 (PUB004). Circular buffer (100 elements).            │
 * │ BOUNDARIES  │ Sample count saturates at windowSize.                               │
 * │             │ Zero-value behavior: valid input, included in average per PUB001.   │
 * ├─────────────┼────────────────────────────────────────────────────────────────────┤
 * │ CITATIONS   │ PUB001: Moving arithmetic mean definition.                          │
 * │             │ PUB002: cyclicExecution periodic update.                            │
 * │             │ PUB003: External trigger rising edge.                               │
 * │             │ PUB004: Reset signal and window validation.                         │
 * │             │ PUB006: 16#0000 success status.                                     │
 * │             │ PUB007: 16#8200 window length error status.                         │
 * └─────────────┴────────────────────────────────────────────────────────────────────┘
 *)
VAR_INPUT
    cyclicExecution : BOOL;
    trigger : BOOL;
    value : LREAL;
    windowSize : INT;
    reset : BOOL;
END_VAR

VAR_OUTPUT
    average : LREAL;
    windowSizeReached : BOOL;
    error : BOOL;
    status : WORD;
END_VAR

VAR
    dataBuffer : ARRAY[1..100] OF LREAL;
    sampleCount : INT := 0;
    sumAccumulator : LREAL := 0.0;
    bufferIndex : INT := 0;
    triggerRisingEdge : BOOL := FALSE;
    prevTrigger : BOOL := FALSE;
END_VAR

IF reset THEN
    sampleCount := 0;
    sumAccumulator := 0.0;
    bufferIndex := 0;
    windowSizeReached := FALSE;
    error := FALSE;
    status := 16#0000;
    triggerRisingEdge := FALSE;
    prevTrigger := FALSE;
END_IF;

IF NOT error AND (cyclicExecution OR triggerRisingEdge) THEN
    bufferIndex := (bufferIndex MOD INT_TO_INT(windowSize)) + 1;

    IF sampleCount >= windowSize THEN
        sumAccumulator := sumAccumulator - dataBuffer[bufferIndex];
    ELSE
        sampleCount := sampleCount + 1;
    END_IF;

    dataBuffer[bufferIndex] := value;
    sumAccumulator := sumAccumulator + value;
    average := sumAccumulator / LREAL_TO_LREAL(INT_TO_LREAL(sampleCount));
    windowSizeReached := (sampleCount >= windowSize);
END_IF;

IF windowSize < 1 OR windowSize > 100 THEN
    error := TRUE;
    status := 16#8200;
END_IF;

prevTrigger := trigger;
triggerRisingEdge := trigger AND NOT prevTrigger;

END_FUNCTION_BLOCK

(* ---- public-medium-03.candidate_02.st ---- *)
FUNCTION_BLOCK FB_MovingAverage
(* Engineering Contract
 * ┌─────────────────────────────────────────────────────────────────────────────────────┐
 * │ OUTPUT STATE TABLE                                                                │
 * ├─────────────┬────────────────────────────────────────────────────────────────────┤
 * │ average     │ HOLD: Retained between scans; updated when valid sample processed.  │
 * │             │ RETAIN on reset: Returns to 0.0 via sum reset.                      │
 * │ windowSizeReached│ ACTIVE: TRUE when sampleCount >= windowSize (PUB001 window).   │
 * │             │ DEACTIVATION: Set FALSE on reset.                                   │
 * │ error       │ ACTIVE: TRUE when windowSize invalid (<1 or >100).                  │
 * │             │ DEACTIVATION: Set FALSE when reset clears error.                    │
 * │ status      │ RETAIN: 16#8200 when invalid windowSize; 16#0000 otherwise.         │
 * │             │ RESET: Set to 16#0000 on valid reset or valid windowSize.           │
 * ├─────────────┼────────────────────────────────────────────────────────────────────┤
 * │ TRIGGER     │ Rising edge on trigger input (PUB003). Edge detection via           │
 * │             │ triggerRisingEdge state variable. Same-scan priority: cyclicExecution│
 * │             │ checked first per PUB002.                                           │
 * ├─────────────┼────────────────────────────────────────────────────────────────────┤
 * │ WINDOW      │ Bounded 1..100 (PUB004). Circular buffer (100 elements).            │
 * │ BOUNDARIES  │ Sample count saturates at windowSize.                               │
 * │             │ Zero-value behavior: valid input, included in average per PUB001.   │
 * ├─────────────┼────────────────────────────────────────────────────────────────────┤
 * │ CITATIONS   │ PUB001: Moving arithmetic mean definition.                          │
 * │             │ PUB002: cyclicExecution periodic update.                            │
 * │             │ PUB003: External trigger rising edge.                               │
 * │             │ PUB004: Reset signal and window validation.                         │
 * │             │ PUB006: 16#0000 success status.                                     │
 * │             │ PUB007: 16#8200 window length error status.                         │
 * └─────────────┴────────────────────────────────────────────────────────────────────┘
 *)
VAR_INPUT
    cyclicExecution : BOOL;
    trigger : BOOL;
    value : LREAL;
    windowSize : INT;
    reset : BOOL;
END_VAR

VAR_OUTPUT
    average : LREAL;
    windowSizeReached : BOOL;
    error : BOOL;
    status : WORD;
END_VAR

VAR
    dataBuffer : ARRAY[1..100] OF LREAL;
    sampleCount : INT := 0;
    sumAccumulator : LREAL := 0.0;
    bufferIndex : INT := 0;
    triggerRisingEdge : BOOL := FALSE;
    prevTrigger : BOOL := FALSE;
END_VAR

IF reset THEN
    sampleCount := 0;
    sumAccumulator := 0.0;
    bufferIndex := 0;
    windowSizeReached := FALSE;
    error := FALSE;
    status := 16#0000;
    triggerRisingEdge := FALSE;
    prevTrigger := FALSE;
END_IF;

IF windowSize < 1 OR windowSize > 100 THEN
    error := TRUE;
    status := 16#8200;
END_IF;

IF NOT error AND (cyclicExecution OR triggerRisingEdge) THEN
    bufferIndex := (bufferIndex MOD windowSize) + 1;

    IF sampleCount >= windowSize THEN
        sumAccumulator := sumAccumulator - dataBuffer[bufferIndex];
    ELSE
        sampleCount := sampleCount + 1;
    END_IF;

    dataBuffer[bufferIndex] := value;
    sumAccumulator := sumAccumulator + value;
    average := sumAccumulator / INT_TO_LREAL(sampleCount);
    windowSizeReached := (sampleCount >= windowSize);
END_IF;

prevTrigger := trigger;
triggerRisingEdge := trigger AND NOT prevTrigger;

END_FUNCTION_BLOCK

(* ---- public-medium-03.raw_candidate_01.st ---- *)
FUNCTION_BLOCK FB_MovingAverage
(* Engineering Contract
 * ┌─────────────────────────────────────────────────────────────────────────────────────┐
 * │ OUTPUT STATE TABLE                                                                │
 * ├─────────────┬────────────────────────────────────────────────────────────────────┤
 * │ average     │ HOLD: Retained between scans; updated when valid sample processed.  │
 * │             │ RETAIN on reset: Returns to 0.0 via sum reset.                      │
 * │ windowSizeReached│ ACTIVE: TRUE when sampleCount >= windowSize (PUB001 window).   │
 * │             │ DEACTIVATION: Set FALSE on reset.                                   │
 * │ error       │ ACTIVE: TRUE when windowSize invalid (<1 or >100).                  │
 * │             │ DEACTIVATION: Set FALSE when reset clears error.                    │
 * │ status      │ RETAIN: 16#8200 when invalid windowSize; 16#0000 otherwise.         │
 * │             │ RESET: Set to 16#0000 on valid reset or valid windowSize.           │
 * ├─────────────┼────────────────────────────────────────────────────────────────────┤
 * │ TRIGGER     │ Rising edge on trigger input (PUB003). Edge detection via           │
 * │             │ triggerPrev state variable. Same-scan priority: cyclicExecution     │
 * │             │ checked first per PUB002.                                           │
 * ├─────────────┼────────────────────────────────────────────────────────────────────┤
 * │ WINDOW      │ Bounded 1..100 (PUB004). Circular buffer (100 elements).            │
 * │ BOUNDARIES  │ Sample count saturates at windowSize.                               │
 * │             │ Zero-value behavior: valid input, included in average per PUB001.   │
 * ├─────────────┼────────────────────────────────────────────────────────────────────┤
 * │ CITATIONS   │ PUB001: Moving arithmetic mean definition.                          │
 * │             │ PUB002: cyclicExecution periodic update.                            │
 * │             │ PUB003: External trigger rising edge.                               │
 * │             │ PUB004: Reset signal and window validation.                         │
 * │             │ PUB006: 16#0000 success status.                                     │
 * │             │ PUB007: 16#8200 window length error status.                         │
 * └─────────────┴────────────────────────────────────────────────────────────────────┘
 *)
VAR_INPUT
    cyclicExecution : BOOL;
    trigger : BOOL;
    value : LREAL;
    windowSize : INT;
    reset : BOOL;
END_VAR

VAR_OUTPUT
    average : LREAL;
    windowSizeReached : BOOL;
    error : BOOL;
    status : WORD;
END_VAR

VAR
    dataBuffer : ARRAY[1..100] OF LREAL;
    sampleCount : INT := 0;
    sumAccumulator : LREAL := 0.0;
    bufferIndex : INT := 0;
    triggerRisingEdge : BOOL := FALSE;
    prevTrigger : BOOL := FALSE;
END_VAR

IF reset THEN
    sampleCount := 0;
    sumAccumulator := 0.0;
    bufferIndex := 0;
    windowSizeReached := FALSE;
    error := FALSE;
    status := 16#0000;
    triggerRisingEdge := FALSE;
    prevTrigger := FALSE;
END_IF;

IF NOT error AND (cyclicExecution OR triggerRisingEdge) THEN
    bufferIndex := (bufferIndex MOD INT_TO_INT(windowSize)) + 1;

    IF sampleCount >= windowSize THEN
        sumAccumulator := sumAccumulator - dataBuffer[bufferIndex];
    ELSE
        sampleCount := sampleCount + 1;
    END_IF;

    dataBuffer[bufferIndex] := value;
    sumAccumulator := sumAccumulator + value;
    average := sumAccumulator / LREAL_TO_LREAL(INT_TO_LREAL(sampleCount));
    windowSizeReached := (sampleCount >= windowSize);
END_IF;

IF windowSize < 1 OR windowSize > 100 THEN
    error := TRUE;
    status := 16#8200;
END_IF;

prevTrigger := trigger;
triggerRisingEdge := trigger AND NOT prevTrigger;

END_FUNCTION_BLOCK

(* ---- public-medium-03.raw_candidate_02.st ---- *)
FUNCTION_BLOCK FB_MovingAverage
(* Engineering Contract
 * ┌─────────────────────────────────────────────────────────────────────────────────────┐
 * │ OUTPUT STATE TABLE                                                                │
 * ├─────────────┬────────────────────────────────────────────────────────────────────┤
 * │ average     │ HOLD: Retained between scans; updated when valid sample processed.  │
 * │             │ RETAIN on reset: Returns to 0.0 via sum reset.                      │
 * │ windowSizeReached│ ACTIVE: TRUE when sampleCount >= windowSize (PUB001 window).   │
 * │             │ DEACTIVATION: Set FALSE on reset.                                   │
 * │ error       │ ACTIVE: TRUE when windowSize invalid (<1 or >100).                  │
 * │             │ DEACTIVATION: Set FALSE when reset clears error.                    │
 * │ status      │ RETAIN: 16#8200 when invalid windowSize; 16#0000 otherwise.         │
 * │             │ RESET: Set to 16#0000 on valid reset or valid windowSize.           │
 * ├─────────────┼────────────────────────────────────────────────────────────────────┤
 * │ TRIGGER     │ Rising edge on trigger input (PUB003). Edge detection via           │
 * │             │ triggerRisingEdge state variable. Same-scan priority: cyclicExecution│
 * │             │ checked first per PUB002.                                           │
 * ├─────────────┼────────────────────────────────────────────────────────────────────┤
 * │ WINDOW      │ Bounded 1..100 (PUB004). Circular buffer (100 elements).            │
 * │ BOUNDARIES  │ Sample count saturates at windowSize.                               │
 * │             │ Zero-value behavior: valid input, included in average per PUB001.   │
 * ├─────────────┼────────────────────────────────────────────────────────────────────┤
 * │ CITATIONS   │ PUB001: Moving arithmetic mean definition.                          │
 * │             │ PUB002: cyclicExecution periodic update.                            │
 * │             │ PUB003: External trigger rising edge.                               │
 * │             │ PUB004: Reset signal and window validation.                         │
 * │             │ PUB006: 16#0000 success status.                                     │
 * │             │ PUB007: 16#8200 window length error status.                         │
 * └─────────────┴────────────────────────────────────────────────────────────────────┘
 *)
VAR_INPUT
    cyclicExecution : BOOL;
    trigger : BOOL;
    value : LREAL;
    windowSize : INT;
    reset : BOOL;
END_VAR

VAR_OUTPUT
    average : LREAL;
    windowSizeReached : BOOL;
    error : BOOL;
    status : WORD;
END_VAR

VAR
    dataBuffer : ARRAY[1..100] OF LREAL;
    sampleCount : INT := 0;
    sumAccumulator : LREAL := 0.0;
    bufferIndex : INT := 0;
    triggerRisingEdge : BOOL := FALSE;
    prevTrigger : BOOL := FALSE;
END_VAR

IF reset THEN
    sampleCount := 0;
    sumAccumulator := 0.0;
    bufferIndex := 0;
    windowSizeReached := FALSE;
    error := FALSE;
    status := 16#0000;
    triggerRisingEdge := FALSE;
    prevTrigger := FALSE;
END_IF;

IF windowSize < 1 OR windowSize > 100 THEN
    error := TRUE;
    status := 16#8200;
END_IF;

IF NOT error AND (cyclicExecution OR triggerRisingEdge) THEN
    bufferIndex := (bufferIndex MOD windowSize) + 1;

    IF sampleCount >= windowSize THEN
        sumAccumulator := sumAccumulator - dataBuffer[bufferIndex];
    ELSE
        sampleCount := sampleCount + 1;
    END_IF;

    dataBuffer[bufferIndex] := value;
    sumAccumulator := sumAccumulator + value;
    average := sumAccumulator / INT_TO_LREAL(sampleCount);
    windowSizeReached := (sampleCount >= windowSize);
END_IF;

prevTrigger := trigger;
triggerRisingEdge := trigger AND NOT prevTrigger;

END_FUNCTION_BLOCK

(* ---- public-medium-04.candidate_01.st ---- *)
(*
ENGINEERING_CONTRACT - FB_TemperatureControl
=============================================
| State/Output          | Activation            | Retention    | Reset/Deactivation           | Priority     | Units/Boundaries        |
|-----------------------|-----------------------|--------------|-------------------------------|--------------|-------------------------|
| HeaterOutput=TRUE     | Temp<SetTemp AND      | Held while   | Temp>=SetTemp OR SensorFault  | Normal:1     | BOOL                    |
|                       | NOT OverheatProtection| conditions   | OR OverheatTriggered          | Fault:1      |                         |
| OverheatProtection=TRUE| After 5s continuous   | Latched      | After 3s wait, then auto      | Same-scan    | BOOL                    |
|                       | HeaterOutput=TRUE     | (PUB006)     | reset (PUB006)                | w/ heater off|                         |
| HeaterStatus          | Direct mirror of      | Same as      | Same as HeaterOutput          | Same-scan    | BOOL                    |
|                       | HeaterOutput          | HeaterOutput |                               |              |                         |
| SensorFault Handling  | Temp<0 OR Temp>100    | Latched      | Temp back in [0,100] range    | Highest      | 0 <= Temp <= 100 (PUB007)|
|                       |                       |              |                               |              |                         |
| CurrentTemperature    | Assign from input     | Real-time    | None (display only)           | Passive      | REAL, fault=0           |
| SetTempDisplay        | Assign from input     | Real-time    | None (display only)           | Passive      | REAL                    |
==============================================================================================================
PUB001: Function block implementation
PUB002: TemperatureSensorInput reading
PUB003-005: Temperature comparison and heater control
PUB006: Overheat protection with 5s trigger, 3s reset
PUB007: Status indication outputs
PUB008: Sensor fault detection (0-100 range)
*)
FUNCTION_BLOCK FB_TemperatureControl
VAR_INPUT
    TemperatureSensorInput : REAL;
    SetTemperature : REAL;
END_VAR
VAR_OUTPUT
    CurrentTemperature : REAL;
    SetTempDisplay : REAL;
    HeaterStatus : BOOL;
    OverheatProtection : BOOL;
    HeaterOutput : BOOL := FALSE;
END_VAR
VAR
    OverheatTimer : TON;
    ResetTimer : TON;
    HeaterRunTimer : TON;
    SensorFault : BOOL := FALSE;
    OverheatTriggered : BOOL := FALSE;
    HeaterShouldBeOn : BOOL := FALSE;
    HeaterOnDuration : TIME := T#0S;
    LastScanHeaterOn : BOOL := FALSE;
END_VAR

// Sensor fault detection (PUB008)
SensorFault := (TemperatureSensorInput < 0.0) OR (TemperatureSensorInput > 100.0);

// Update displays (PUB007)
CurrentTemperature := TemperatureSensorInput;
SetTempDisplay := SetTemperature;

// Normal temperature control logic (PUB003, PUB004)
// If sensor fault, heater should be off
IF NOT SensorFault THEN
    HeaterShouldBeOn := (TemperatureSensorInput < SetTemperature);
ELSE
    HeaterShouldBeOn := FALSE;
END_IF;

// Overheat protection logic (PUB006)
// Track continuous heater on time
IF HeaterShouldBeOn AND NOT OverheatTriggered THEN
    HeaterOnDuration := HeaterOnDuration + T#1S; // Assuming 1s scan time
    IF HeaterOnDuration >= T#5S THEN
        OverheatTriggered := TRUE;
    END_IF;
ELSE
    HeaterOnDuration := T#0S;
END_IF;

// Handle overheat protection state (PUB006)
IF OverheatTriggered THEN
    OverheatProtection := TRUE;
    HeaterOutput := FALSE;
    // Start 3s reset timer after overheat triggered
    ResetTimer(IN := TRUE, PT := T#3S);
    IF ResetTimer.Q THEN
        OverheatTriggered := FALSE;
        OverheatProtection := FALSE;
        ResetTimer(IN := FALSE);
        ResetTimer();
    END_IF;
ELSE
    ResetTimer(IN := FALSE);
    ResetTimer();
    OverheatProtection := FALSE;
    // Normal operation - heater follows temperature comparison
    HeaterOutput := HeaterShouldBeOn;
END_IF;

// Update heater status display (PUB007)
HeaterStatus := HeaterOutput;

END_FUNCTION_BLOCK

(* ---- public-medium-04.candidate_02.st ---- *)
(*
ENGINEERING_CONTRACT - FB_TemperatureControl
=============================================
| State/Output          | Activation            | Retention    | Reset/Deactivation           | Priority     | Units/Boundaries        |
|-----------------------|-----------------------|--------------|-------------------------------|--------------|-------------------------|
| HeaterOutput=TRUE     | Temp<SetTemp AND      | Held while   | Temp>=SetTemp OR SensorFault  | Normal:1     | BOOL                    |
|                       | NOT OverheatProtection| conditions   | OR OverheatTriggered          | Fault:1      |                         |
| OverheatProtection=TRUE| After 5s continuous   | Latched      | After 3s wait, then auto      | Same-scan    | BOOL                    |
|                       | HeaterOutput=TRUE     | (PUB006)     | reset (PUB006)                | w/ heater off|                         |
| HeaterStatus          | Direct mirror of      | Same as      | Same as HeaterOutput          | Same-scan    | BOOL                    |
|                       | HeaterOutput          | HeaterOutput |                               |              |                         |
| SensorFault Handling  | Temp<0 OR Temp>100    | Latched      | Temp back in [0,100] range    | Highest      | 0 <= Temp <= 100 (PUB007)|
|                       |                       |              |                               |              |                         |
| CurrentTemperature    | Assign from input     | Real-time    | None (display only)           | Passive      | REAL, fault=0           |
| SetTempDisplay        | Assign from input     | Real-time    | None (display only)           | Passive      | REAL                    |
==============================================================================================================
PUB001: Function block implementation
PUB002: TemperatureSensorInput reading
PUB003-005: Temperature comparison and heater control
PUB006: Overheat protection with 5s trigger, 3s reset
PUB007: Status indication outputs
PUB008: Sensor fault detection (0-100 range)
*)
FUNCTION_BLOCK FB_TemperatureControl
VAR_INPUT
    TemperatureSensorInput : REAL;
    SetTemperature : REAL;
END_VAR
VAR_OUTPUT
    CurrentTemperature : REAL;
    SetTempDisplay : REAL;
    HeaterStatus : BOOL;
    OverheatProtection : BOOL;
    HeaterOutput : BOOL := FALSE;
END_VAR
VAR
    tonOverheat : TON;
    tonReset : TON;
    SensorFault : BOOL := FALSE;
    OverheatTriggered : BOOL := FALSE;
END_VAR

// Sensor fault detection (PUB008)
SensorFault := (TemperatureSensorInput < 0.0) OR (TemperatureSensorInput > 100.0);

// Update displays (PUB007)
CurrentTemperature := TemperatureSensorInput;
SetTempDisplay := SetTemperature;

// Overheat protection logic (PUB006)
IF OverheatTriggered THEN
    // Overheat active - heater off, start reset timer
    OverheatProtection := TRUE;
    HeaterOutput := FALSE;
    tonOverheat(IN := FALSE);
    tonOverheat();
    tonReset(IN := TRUE, PT := T#3S);
    IF tonReset.Q THEN
        OverheatTriggered := FALSE;
        OverheatProtection := FALSE;
        tonReset(IN := FALSE);
        tonReset();
    END_IF;
ELSE
    // Normal operation
    tonReset(IN := FALSE);
    tonReset();
    OverheatProtection := FALSE;

    // Start overheat timer when heater would be on
    IF NOT SensorFault AND (TemperatureSensorInput < SetTemperature) THEN
        tonOverheat(IN := TRUE, PT := T#5S);
    ELSE
        tonOverheat(IN := FALSE);
    END_IF;
    tonOverheat();

    // Check if overheat threshold reached
    IF tonOverheat.Q THEN
        OverheatTriggered := TRUE;
        HeaterOutput := FALSE;
    ELSE
        // Normal heater control (PUB003, PUB004, PUB005)
        IF NOT SensorFault THEN
            IF TemperatureSensorInput < SetTemperature THEN
                HeaterOutput := TRUE;
            ELSE
                HeaterOutput := FALSE;
            END_IF;
        ELSE
            HeaterOutput := FALSE;
        END_IF;
    END_IF;
END_IF;

// Update heater status display (PUB007)
HeaterStatus := HeaterOutput;

END_FUNCTION_BLOCK

(* ---- public-medium-04.raw_candidate_01.st ---- *)
(*
ENGINEERING_CONTRACT - FB_TemperatureControl
=============================================
| State/Output          | Activation            | Retention    | Reset/Deactivation           | Priority     | Units/Boundaries        |
|-----------------------|-----------------------|--------------|-------------------------------|--------------|-------------------------|
| HeaterOutput=TRUE     | Temp<SetTemp AND      | Held while   | Temp>=SetTemp OR SensorFault  | Normal:1     | BOOL                    |
|                       | NOT OverheatProtection| conditions   | OR OverheatTriggered          | Fault:1      |                         |
| OverheatProtection=TRUE| After 5s continuous   | Latched      | After 3s wait, then auto      | Same-scan    | BOOL                    |
|                       | HeaterOutput=TRUE     | (PUB006)     | reset (PUB006)                | w/ heater off|                         |
| HeaterStatus          | Direct mirror of      | Same as      | Same as HeaterOutput          | Same-scan    | BOOL                    |
|                       | HeaterOutput          | HeaterOutput |                               |              |                         |
| SensorFault Handling  | Temp<0 OR Temp>100    | Latched      | Temp back in [0,100] range    | Highest      | 0 <= Temp <= 100 (PUB007)|
|                       |                       |              |                               |              |                         |
| CurrentTemperature    | Assign from input     | Real-time    | None (display only)           | Passive      | REAL, fault=0           |
| SetTempDisplay        | Assign from input     | Real-time    | None (display only)           | Passive      | REAL                    |
==============================================================================================================
PUB001: Function block implementation
PUB002: TemperatureSensorInput reading
PUB003-005: Temperature comparison and heater control
PUB006: Overheat protection with 5s trigger, 3s reset
PUB007: Status indication outputs
PUB008: Sensor fault detection (0-100 range)
*)
FUNCTION_BLOCK FB_TemperatureControl
VAR_INPUT
    TemperatureSensorInput : REAL;
    SetTemperature : REAL;
END_VAR
VAR_OUTPUT
    CurrentTemperature : REAL;
    SetTempDisplay : REAL;
    HeaterStatus : BOOL;
    OverheatProtection : BOOL;
    HeaterOutput : BOOL := FALSE;
END_VAR
VAR
    OverheatTimer : TON;
    ResetTimer : TON;
    HeaterRunTimer : TON;
    SensorFault : BOOL := FALSE;
    OverheatTriggered : BOOL := FALSE;
    HeaterShouldBeOn : BOOL := FALSE;
    HeaterOnDuration : TIME := T#0S;
    LastScanHeaterOn : BOOL := FALSE;
END_VAR

// Sensor fault detection (PUB008)
SensorFault := (TemperatureSensorInput < 0.0) OR (TemperatureSensorInput > 100.0);

// Update displays (PUB007)
CurrentTemperature := TemperatureSensorInput;
SetTempDisplay := SetTemperature;

// Normal temperature control logic (PUB003, PUB004)
// If sensor fault, heater should be off
IF NOT SensorFault THEN
    HeaterShouldBeOn := (TemperatureSensorInput < SetTemperature);
ELSE
    HeaterShouldBeOn := FALSE;
END_IF;

// Overheat protection logic (PUB006)
// Track continuous heater on time
IF HeaterShouldBeOn AND NOT OverheatTriggered THEN
    HeaterOnDuration := HeaterOnDuration + T#1S; // Assuming 1s scan time
    IF HeaterOnDuration >= T#5S THEN
        OverheatTriggered := TRUE;
    END_IF;
ELSE
    HeaterOnDuration := T#0S;
END_IF;

// Handle overheat protection state (PUB006)
IF OverheatTriggered THEN
    OverheatProtection := TRUE;
    HeaterOutput := FALSE;
    // Start 3s reset timer after overheat triggered
    ResetTimer(IN := TRUE, PT := T#3S);
    IF ResetTimer.Q THEN
        OverheatTriggered := FALSE;
        OverheatProtection := FALSE;
        ResetTimer(IN := FALSE);
        ResetTimer();
    END_IF;
ELSE
    ResetTimer(IN := FALSE);
    ResetTimer();
    OverheatProtection := FALSE;
    // Normal operation - heater follows temperature comparison
    HeaterOutput := HeaterShouldBeOn;
END_IF;

// Update heater status display (PUB007)
HeaterStatus := HeaterOutput;

END_FUNCTION_BLOCK

(* ---- public-medium-04.raw_candidate_02.st ---- *)
(*
ENGINEERING_CONTRACT - FB_TemperatureControl
=============================================
| State/Output          | Activation            | Retention    | Reset/Deactivation           | Priority     | Units/Boundaries        |
|-----------------------|-----------------------|--------------|-------------------------------|--------------|-------------------------|
| HeaterOutput=TRUE     | Temp<SetTemp AND      | Held while   | Temp>=SetTemp OR SensorFault  | Normal:1     | BOOL                    |
|                       | NOT OverheatProtection| conditions   | OR OverheatTriggered          | Fault:1      |                         |
| OverheatProtection=TRUE| After 5s continuous   | Latched      | After 3s wait, then auto      | Same-scan    | BOOL                    |
|                       | HeaterOutput=TRUE     | (PUB006)     | reset (PUB006)                | w/ heater off|                         |
| HeaterStatus          | Direct mirror of      | Same as      | Same as HeaterOutput          | Same-scan    | BOOL                    |
|                       | HeaterOutput          | HeaterOutput |                               |              |                         |
| SensorFault Handling  | Temp<0 OR Temp>100    | Latched      | Temp back in [0,100] range    | Highest      | 0 <= Temp <= 100 (PUB007)|
|                       |                       |              |                               |              |                         |
| CurrentTemperature    | Assign from input     | Real-time    | None (display only)           | Passive      | REAL, fault=0           |
| SetTempDisplay        | Assign from input     | Real-time    | None (display only)           | Passive      | REAL                    |
==============================================================================================================
PUB001: Function block implementation
PUB002: TemperatureSensorInput reading
PUB003-005: Temperature comparison and heater control
PUB006: Overheat protection with 5s trigger, 3s reset
PUB007: Status indication outputs
PUB008: Sensor fault detection (0-100 range)
*)
FUNCTION_BLOCK FB_TemperatureControl
VAR_INPUT
    TemperatureSensorInput : REAL;
    SetTemperature : REAL;
END_VAR
VAR_OUTPUT
    CurrentTemperature : REAL;
    SetTempDisplay : REAL;
    HeaterStatus : BOOL;
    OverheatProtection : BOOL;
    HeaterOutput : BOOL := FALSE;
END_VAR
VAR
    tonOverheat : TON;
    tonReset : TON;
    SensorFault : BOOL := FALSE;
    OverheatTriggered : BOOL := FALSE;
END_VAR

// Sensor fault detection (PUB008)
SensorFault := (TemperatureSensorInput < 0.0) OR (TemperatureSensorInput > 100.0);

// Update displays (PUB007)
CurrentTemperature := TemperatureSensorInput;
SetTempDisplay := SetTemperature;

// Overheat protection logic (PUB006)
IF OverheatTriggered THEN
    // Overheat active - heater off, start reset timer
    OverheatProtection := TRUE;
    HeaterOutput := FALSE;
    tonOverheat(IN := FALSE);
    tonOverheat();
    tonReset(IN := TRUE, PT := T#3S);
    IF tonReset.Q THEN
        OverheatTriggered := FALSE;
        OverheatProtection := FALSE;
        tonReset(IN := FALSE);
        tonReset();
    END_IF;
ELSE
    // Normal operation
    tonReset(IN := FALSE);
    tonReset();
    OverheatProtection := FALSE;

    // Start overheat timer when heater would be on
    IF NOT SensorFault AND (TemperatureSensorInput < SetTemperature) THEN
        tonOverheat(IN := TRUE, PT := T#5S);
    ELSE
        tonOverheat(IN := FALSE);
    END_IF;
    tonOverheat();

    // Check if overheat threshold reached
    IF tonOverheat.Q THEN
        OverheatTriggered := TRUE;
        HeaterOutput := FALSE;
    ELSE
        // Normal heater control (PUB003, PUB004, PUB005)
        IF NOT SensorFault THEN
            IF TemperatureSensorInput < SetTemperature THEN
                HeaterOutput := TRUE;
            ELSE
                HeaterOutput := FALSE;
            END_IF;
        ELSE
            HeaterOutput := FALSE;
        END_IF;
    END_IF;
END_IF;

// Update heater status display (PUB007)
HeaterStatus := HeaterOutput;

END_FUNCTION_BLOCK

(* ---- public-medium-08.candidate_01.st ---- *)
FUNCTION_BLOCK IPv4_Parser
(*
ENGINEERING_CONTRACT
===================
PUB001-003: Parse dotted-decimal IPv4 string to 32-bit UDINT in network byte order
PUB004:     Output = 0 for invalid input (incl. valid 0.0.0.0 → ambiguity resolved as 0)

OUTPUT STATE:
- ipValue: activation = parsed value, retention = n/a, reset = n/a (one-shot per call)
- Units: 0–4294967295 (32-bit), zero on any malformed input per PUB004

VALIDATION (in priority order):
1. Exactly three dot separators found, each at valid position
2. No fourth dot after third (prevents extra segments)
3. Four nonempty segments, each 1–3 chars
4. Each segment contains only decimal digits (char '0'–'9')
5. Each segment numeric value within 0–255

ASSEMBLY: Network byte order per PUB003
- Segment 1 → bits[31:24] (MSB)
- Segment 2 → bits[23:16]
- Segment 3 → bits[15:8]
- Segment 4 → bits[7:0] (LSB)

SCAN BEHAVIOR: Deterministic single-scan parse, no latching, no edge triggers
*)

VAR_INPUT
    ipText : STRING(254);
END_VAR

VAR_OUTPUT
    ipValue : UDINT := 0;
END_VAR

VAR
    dotPos1   : INT;
    dotPos2   : INT;
    dotPos3   : INT;
    textLen   : INT;
    segLen    : INT;
    seg1      : STRING(3);
    seg2      : STRING(3);
    seg3      : STRING(3);
    seg4      : STRING(3);
    val1      : UDINT;
    val2      : UDINT;
    val3      : UDINT;
    val4      : UDINT;
    i         : INT;
    charVal   : BYTE;
    valid     : BOOL;
END_VAR

    // Locate the three period separators
    dotPos1 := FIND(ipText, '.');
    dotPos2 := FIND(ipText, '.', dotPos1 + 1);
    dotPos3 := FIND(ipText, '.', dotPos2 + 1);

    // PUB002: must have exactly three dots at valid positions
    IF dotPos1 <= 0 OR dotPos2 <= 0 OR dotPos3 <= 0 THEN
        ipValue := 0;
        RETURN;
    END_IF;

    // No fourth dot allowed
    textLen := LEN(ipText);
    IF FIND(ipText, '.', dotPos3 + 1) <> 0 THEN
        ipValue := 0;
        RETURN;
    END_IF;

    // Segment 1: positions 1 to dotPos1-1 (length = dotPos1-1)
    segLen := dotPos1 - 1;
    IF segLen < 1 OR segLen > 3 THEN
        ipValue := 0;
        RETURN;
    END_IF;
    seg1 := MID(ipText, segLen, 1);
    valid := TRUE;
    FOR i := 1 TO segLen DO
        charVal := TO_BYTE(MID(seg1, 1, i));
        IF charVal < 48 OR charVal > 57 THEN
            valid := FALSE;
            EXIT;
        END_IF;
    END_FOR;
    IF NOT valid THEN
        ipValue := 0;
        RETURN;
    END_IF;
    val1 := TO_UDINT(seg1);
    IF val1 > 255 THEN
        ipValue := 0;
        RETURN;
    END_IF;

    // Segment 2: positions dotPos1+1 to dotPos2-1
    segLen := dotPos2 - dotPos1 - 1;
    IF segLen < 1 OR segLen > 3 THEN
        ipValue := 0;
        RETURN;
    END_IF;
    seg2 := MID(ipText, segLen, dotPos1 + 1);
    valid := TRUE;
    FOR i := 1 TO segLen DO
        charVal := TO_BYTE(MID(seg2, 1, i));
        IF charVal < 48 OR charVal > 57 THEN
            valid := FALSE;
            EXIT;
        END_IF;
    END_FOR;
    IF NOT valid THEN
        ipValue := 0;
        RETURN;
    END_IF;
    val2 := TO_UDINT(seg2);
    IF val2 > 255 THEN
        ipValue := 0;
        RETURN;
    END_IF;

    // Segment 3: positions dotPos2+1 to dotPos3-1
    segLen := dotPos3 - dotPos2 - 1;
    IF segLen < 1 OR segLen > 3 THEN
        ipValue := 0;
        RETURN;
    END_IF;
    seg3 := MID(ipText, segLen, dotPos2 + 1);
    valid := TRUE;
    FOR i := 1 TO segLen DO
        charVal := TO_BYTE(MID(seg3, 1, i));
        IF charVal < 48 OR charVal > 57 THEN
            valid := FALSE;
            EXIT;
        END_IF;
    END_FOR;
    IF NOT valid THEN
        ipValue := 0;
        RETURN;
    END_IF;
    val3 := TO_UDINT(seg3);
    IF val3 > 255 THEN
        ipValue := 0;
        RETURN;
    END_IF;

    // Segment 4: positions dotPos3+1 to end
    segLen := textLen - dotPos3;
    IF segLen < 1 OR segLen > 3 THEN
        ipValue := 0;
        RETURN;
    END_IF;
    seg4 := MID(ipText, segLen, dotPos3 + 1);
    valid := TRUE;
    FOR i := 1 TO segLen DO
        charVal := TO_BYTE(MID(seg4, 1, i));
        IF charVal < 48 OR charVal > 57 THEN
            valid := FALSE;
            EXIT;
        END_IF;
    END_FOR;
    IF NOT valid THEN
        ipValue := 0;
        RETURN;
    END_IF;
    val4 := TO_UDINT(seg4);
    IF val4 > 255 THEN
        ipValue := 0;
        RETURN;
    END_IF;

    // PUB003: Assemble in network byte order (MSB first)
    ipValue := SHL(val1, 24) OR SHL(val2, 16) OR SHL(val3, 8) OR val4;

END_FUNCTION_BLOCK

(* ---- public-medium-08.candidate_02.st ---- *)
FUNCTION_BLOCK IPv4_Parser
(*
ENGINEERING_CONTRACT
===================
PUB001-003: Parse dotted-decimal IPv4 string to 32-bit UDINT in network byte order
PUB004:     Output = 0 for invalid input (incl. valid 0.0.0.0 → ambiguity resolved as 0)

OUTPUT STATE:
- ipValue: activation = parsed value, retention = n/a, reset = n/a (one-shot per call)
- Units: 0–4294967295 (32-bit), zero on any malformed input per PUB004

VALIDATION (in priority order):
1. Exactly three dot separators found, each at valid position
2. No fourth dot after third (prevents extra segments)
3. Four nonempty segments, each 1–3 chars
4. Each segment contains only decimal digits (char '0'–'9')
5. Each segment numeric value within 0–255

ASSEMBLY: Network byte order per PUB003
- Segment 1 → bits[31:24] (MSB)
- Segment 2 → bits[23:16]
- Segment 3 → bits[15:8]
- Segment 4 → bits[7:0] (LSB)

SCAN BEHAVIOR: Deterministic single-scan parse, no latching, no edge triggers
*)

VAR_INPUT
    ipText : STRING(254);
END_VAR

VAR_OUTPUT
    ipValue : UDINT := 0;
END_VAR

VAR
    dotPos1   : INT;
    dotPos2   : INT;
    dotPos3   : INT;
    textLen   : INT;
    segLen    : INT;
    seg1      : STRING(3);
    seg2      : STRING(3);
    seg3      : STRING(3);
    seg4      : STRING(3);
    val1      : UDINT;
    val2      : UDINT;
    val3      : UDINT;
    val4      : UDINT;
    i         : INT;
    charVal   : BYTE;
    valid     : BOOL;
    remainder : STRING(254);
END_VAR

    textLen := LEN(ipText);

    // Locate the three period separators using substring search (FIND takes 2 args only)
    dotPos1 := FIND(ipText, '.');
    IF dotPos1 <= 0 THEN
        ipValue := 0;
        RETURN;
    END_IF;

    remainder := MID(ipText, textLen - dotPos1, dotPos1 + 1);
    dotPos2 := dotPos1 + 1 + FIND(remainder, '.');
    IF dotPos2 <= dotPos1 THEN
        ipValue := 0;
        RETURN;
    END_IF;

    remainder := MID(ipText, textLen - dotPos2, dotPos2 + 1);
    dotPos3 := dotPos2 + 1 + FIND(remainder, '.');
    IF dotPos3 <= dotPos2 THEN
        ipValue := 0;
        RETURN;
    END_IF;

    // No fourth dot allowed
    remainder := MID(ipText, textLen - dotPos3, dotPos3 + 1);
    IF FIND(remainder, '.') > 0 THEN
        ipValue := 0;
        RETURN;
    END_IF;

    // Segment 1: positions 1 to dotPos1-1 (length = dotPos1-1)
    segLen := dotPos1 - 1;
    IF segLen < 1 OR segLen > 3 THEN
        ipValue := 0;
        RETURN;
    END_IF;
    seg1 := MID(ipText, segLen, 1);
    valid := TRUE;
    FOR i := 1 TO segLen DO
        charVal := TO_BYTE(MID(seg1, 1, i));
        IF charVal < 48 OR charVal > 57 THEN
            valid := FALSE;
            EXIT;
        END_IF;
    END_FOR;
    IF NOT valid THEN
        ipValue := 0;
        RETURN;
    END_IF;
    val1 := TO_UDINT(seg1);
    IF val1 > 255 THEN
        ipValue := 0;
        RETURN;
    END_IF;

    // Segment 2: positions dotPos1+1 to dotPos2-1
    segLen := dotPos2 - dotPos1 - 1;
    IF segLen < 1 OR segLen > 3 THEN
        ipValue := 0;
        RETURN;
    END_IF;
    seg2 := MID(ipText, segLen, dotPos1 + 1);
    valid := TRUE;
    FOR i := 1 TO segLen DO
        charVal := TO_BYTE(MID(seg2, 1, i));
        IF charVal < 48 OR charVal > 57 THEN
            valid := FALSE;
            EXIT;
        END_IF;
    END_FOR;
    IF NOT valid THEN
        ipValue := 0;
        RETURN;
    END_IF;
    val2 := TO_UDINT(seg2);
    IF val2 > 255 THEN
        ipValue := 0;
        RETURN;
    END_IF;

    // Segment 3: positions dotPos2+1 to dotPos3-1
    segLen := dotPos3 - dotPos2 - 1;
    IF segLen < 1 OR segLen > 3 THEN
        ipValue := 0;
        RETURN;
    END_IF;
    seg3 := MID(ipText, segLen, dotPos2 + 1);
    valid := TRUE;
    FOR i := 1 TO segLen DO
        charVal := TO_BYTE(MID(seg3, 1, i));
        IF charVal < 48 OR charVal > 57 THEN
            valid := FALSE;
            EXIT;
        END_IF;
    END_FOR;
    IF NOT valid THEN
        ipValue := 0;
        RETURN;
    END_IF;
    val3 := TO_UDINT(seg3);
    IF val3 > 255 THEN
        ipValue := 0;
        RETURN;
    END_IF;

    // Segment 4: positions dotPos3+1 to end
    segLen := textLen - dotPos3;
    IF segLen < 1 OR segLen > 3 THEN
        ipValue := 0;
        RETURN;
    END_IF;
    seg4 := MID(ipText, segLen, dotPos3 + 1);
    valid := TRUE;
    FOR i := 1 TO segLen DO
        charVal := TO_BYTE(MID(seg4, 1, i));
        IF charVal < 48 OR charVal > 57 THEN
            valid := FALSE;
            EXIT;
        END_IF;
    END_FOR;
    IF NOT valid THEN
        ipValue := 0;
        RETURN;
    END_IF;
    val4 := TO_UDINT(seg4);
    IF val4 > 255 THEN
        ipValue := 0;
        RETURN;
    END_IF;

    // PUB003: Assemble in network byte order (MSB first)
    ipValue := SHL(val1, 24) OR SHL(val2, 16) OR SHL(val3, 8) OR val4;

END_FUNCTION_BLOCK

(* ---- public-medium-08.raw_candidate_01.st ---- *)
FUNCTION_BLOCK IPv4_Parser
(*
ENGINEERING_CONTRACT
===================
PUB001-003: Parse dotted-decimal IPv4 string to 32-bit UDINT in network byte order
PUB004:     Output = 0 for invalid input (incl. valid 0.0.0.0 → ambiguity resolved as 0)

OUTPUT STATE:
- ipValue: activation = parsed value, retention = n/a, reset = n/a (one-shot per call)
- Units: 0–4294967295 (32-bit), zero on any malformed input per PUB004

VALIDATION (in priority order):
1. Exactly three dot separators found, each at valid position
2. No fourth dot after third (prevents extra segments)
3. Four nonempty segments, each 1–3 chars
4. Each segment contains only decimal digits (char '0'–'9')
5. Each segment numeric value within 0–255

ASSEMBLY: Network byte order per PUB003
- Segment 1 → bits[31:24] (MSB)
- Segment 2 → bits[23:16]
- Segment 3 → bits[15:8]
- Segment 4 → bits[7:0] (LSB)

SCAN BEHAVIOR: Deterministic single-scan parse, no latching, no edge triggers
*)

VAR_INPUT
    ipText : STRING(254);
END_VAR

VAR_OUTPUT
    ipValue : UDINT := 0;
END_VAR

VAR
    dotPos1   : INT;
    dotPos2   : INT;
    dotPos3   : INT;
    textLen   : INT;
    segLen    : INT;
    seg1      : STRING(3);
    seg2      : STRING(3);
    seg3      : STRING(3);
    seg4      : STRING(3);
    val1      : UDINT;
    val2      : UDINT;
    val3      : UDINT;
    val4      : UDINT;
    i         : INT;
    charVal   : BYTE;
    valid     : BOOL;
END_VAR

    // Locate the three period separators
    dotPos1 := FIND(ipText, '.');
    dotPos2 := FIND(ipText, '.', dotPos1 + 1);
    dotPos3 := FIND(ipText, '.', dotPos2 + 1);

    // PUB002: must have exactly three dots at valid positions
    IF dotPos1 <= 0 OR dotPos2 <= 0 OR dotPos3 <= 0 THEN
        ipValue := 0;
        RETURN;
    END_IF;

    // No fourth dot allowed
    textLen := LEN(ipText);
    IF FIND(ipText, '.', dotPos3 + 1) <> 0 THEN
        ipValue := 0;
        RETURN;
    END_IF;

    // Segment 1: positions 1 to dotPos1-1 (length = dotPos1-1)
    segLen := dotPos1 - 1;
    IF segLen < 1 OR segLen > 3 THEN
        ipValue := 0;
        RETURN;
    END_IF;
    seg1 := MID(ipText, segLen, 1);
    valid := TRUE;
    FOR i := 1 TO segLen DO
        charVal := TO_BYTE(MID(seg1, 1, i));
        IF charVal < 48 OR charVal > 57 THEN
            valid := FALSE;
            EXIT;
        END_IF;
    END_FOR;
    IF NOT valid THEN
        ipValue := 0;
        RETURN;
    END_IF;
    val1 := TO_UDINT(seg1);
    IF val1 > 255 THEN
        ipValue := 0;
        RETURN;
    END_IF;

    // Segment 2: positions dotPos1+1 to dotPos2-1
    segLen := dotPos2 - dotPos1 - 1;
    IF segLen < 1 OR segLen > 3 THEN
        ipValue := 0;
        RETURN;
    END_IF;
    seg2 := MID(ipText, segLen, dotPos1 + 1);
    valid := TRUE;
    FOR i := 1 TO segLen DO
        charVal := TO_BYTE(MID(seg2, 1, i));
        IF charVal < 48 OR charVal > 57 THEN
            valid := FALSE;
            EXIT;
        END_IF;
    END_FOR;
    IF NOT valid THEN
        ipValue := 0;
        RETURN;
    END_IF;
    val2 := TO_UDINT(seg2);
    IF val2 > 255 THEN
        ipValue := 0;
        RETURN;
    END_IF;

    // Segment 3: positions dotPos2+1 to dotPos3-1
    segLen := dotPos3 - dotPos2 - 1;
    IF segLen < 1 OR segLen > 3 THEN
        ipValue := 0;
        RETURN;
    END_IF;
    seg3 := MID(ipText, segLen, dotPos2 + 1);
    valid := TRUE;
    FOR i := 1 TO segLen DO
        charVal := TO_BYTE(MID(seg3, 1, i));
        IF charVal < 48 OR charVal > 57 THEN
            valid := FALSE;
            EXIT;
        END_IF;
    END_FOR;
    IF NOT valid THEN
        ipValue := 0;
        RETURN;
    END_IF;
    val3 := TO_UDINT(seg3);
    IF val3 > 255 THEN
        ipValue := 0;
        RETURN;
    END_IF;

    // Segment 4: positions dotPos3+1 to end
    segLen := textLen - dotPos3;
    IF segLen < 1 OR segLen > 3 THEN
        ipValue := 0;
        RETURN;
    END_IF;
    seg4 := MID(ipText, segLen, dotPos3 + 1);
    valid := TRUE;
    FOR i := 1 TO segLen DO
        charVal := TO_BYTE(MID(seg4, 1, i));
        IF charVal < 48 OR charVal > 57 THEN
            valid := FALSE;
            EXIT;
        END_IF;
    END_FOR;
    IF NOT valid THEN
        ipValue := 0;
        RETURN;
    END_IF;
    val4 := TO_UDINT(seg4);
    IF val4 > 255 THEN
        ipValue := 0;
        RETURN;
    END_IF;

    // PUB003: Assemble in network byte order (MSB first)
    ipValue := SHL(val1, 24) OR SHL(val2, 16) OR SHL(val3, 8) OR val4;

END_FUNCTION_BLOCK
